// TIA Portal V21 export
// export: Created 2026-11-07T15:25:00.5686842Z, ExportSetting WithDefaults, DisplayName Totally Integrated Automation Portal, DisplayVersion V21, DisplayName STEP 7 Professional, DisplayVersion V21, DisplayName STEP 7 Safety, DisplayVersion V21, DisplayName Tech WebApplication, DisplayVersion V21, DisplayName WinCC Basic/Comfort/Advanced, DisplayVersion V21, DisplayName WinCC Unified, DisplayVersion V21
Screen "R10_LampA"  1024x768, Number=50, Template=Tpl
  ScreenLayer 
    Rectangle "P_LampAlarm" at 10,10 size 100x30  StyleItem=Rectangle
      RangeAppearanceAnimation "RangeAppearanceAnimation"
        tag P_SwOn
        0..0: back #aaaaaa, fore #000000
        1..1: back #dc0000, fore #000000, flashing
